// TwinCAT 3 PLC project MyLibrary_Test
// ProgramVersion: 3.1.4023.0
// libraries:
//   MyLibrary, * (FabioBolognesi)
//   TcUnit, * (www.tcunit.org)
//   Tc2_Standard, * (Beckhoff Automation GmbH)
//   Tc2_System, * (Beckhoff Automation GmbH)
//   Tc3_Module, * (Beckhoff Automation GmbH)
// project tree:
//   / PlcTask.TcTTO
//   PROGRAMs/ MAIN.TcPOU
//   TESTs/ FB_Conversion_Test.TcPOU, FB_Interpolate_Test.TcPOU, FB_Math_Test.TcPOU, FB_StringBuilder_Test.TcPOU, FB_Sweep_Test.TcPOU, FB_Timer_Test.TcPOU

CONFIGURATION MyLibrary_Test
    RESOURCE PLC ON TwinCAT3
        TASK PlcTask(INTERVAL := T#10ms, PRIORITY := 20);
        PROGRAM MAIN WITH PlcTask : MAIN;
    END_RESOURCE
END_CONFIGURATION

// ---- PROGRAMs/MAIN.TcPOU
// PROGRAMMA DEI TEST: basta dichiarare un'istanza di ogni test suite e chiamare TcUnit.RUN().
// Per aggiungere una suite: crearla in TESTs (EXTENDS TcUnit.FB_TestSuite) e dichiararla qui.
PROGRAM MAIN
VAR
	fbInterpolateTest		:	FB_Interpolate_Test;
	fbMathTest				:	FB_Math_Test;
	fbConversionTest		:	FB_Conversion_Test;
	fbTimerTest				:	FB_Timer_Test;
	fbSweepTest				:	FB_Sweep_Test;
	fbStringBuilderTest		:	FB_StringBuilder_Test;
END_VAR

TcUnit.RUN();

END_PROGRAM

// ---- TESTs/FB_Interpolate_Test.TcPOU
// TEST DI F_InterpolateReal E F_InterpolateTime
FUNCTION_BLOCK FB_Interpolate_Test EXTENDS TcUnit.FB_TestSuite
VAR
END_VAR

MidPoint();
ClampBelow();
ClampAbove();
ReversedPoints();
SamePoints();
InterpolateTime();

METHOD PRIVATE ClampAbove
TEST('ClampAbove');

AssertEquals_REAL(
	Expected	:=	100,
	Actual		:=	ML.F_InterpolateReal(rX0 := 0, rX1 := 10, rY0 := 0, rY1 := 100, rX := 20),
	Delta		:=	0.0001,
	Message		:=	'Dopo il secondo punto deve restituire rY1');

TEST_FINISHED();
END_METHOD

METHOD PRIVATE ClampBelow
TEST('ClampBelow');

AssertEquals_REAL(
	Expected	:=	0,
	Actual		:=	ML.F_InterpolateReal(rX0 := 0, rX1 := 10, rY0 := 0, rY1 := 100, rX := -5),
	Delta		:=	0.0001,
	Message		:=	'Prima del primo punto deve restituire rY0');

TEST_FINISHED();
END_METHOD

METHOD PRIVATE InterpolateTime
TEST('InterpolateTime');

AssertEquals_REAL(
	Expected	:=	2.5,
	Actual		:=	ML.F_InterpolateTime(tX0 := T#0S, tX1 := T#2S, rY0 := 0, rY1 := 10, tX := T#500MS),
	Delta		:=	0.0001,
	Message		:=	'Interpolazione con ascisse TIME');

TEST_FINISHED();
END_METHOD

METHOD PRIVATE MidPoint
TEST('MidPoint');

AssertEquals_REAL(
	Expected	:=	50,
	Actual		:=	ML.F_InterpolateReal(rX0 := 0, rX1 := 10, rY0 := 0, rY1 := 100, rX := 5),
	Delta		:=	0.0001,
	Message		:=	'Punto medio');

TEST_FINISHED();
END_METHOD

METHOD PRIVATE ReversedPoints
TEST('ReversedPoints');

AssertEquals_REAL(
	Expected	:=	25,
	Actual		:=	ML.F_InterpolateReal(rX0 := 10, rX1 := 0, rY0 := 100, rY1 := 0, rX := 2.5),
	Delta		:=	0.0001,
	Message		:=	'Punti in ordine decrescente: interpolazione');
AssertEquals_REAL(
	Expected	:=	100,
	Actual		:=	ML.F_InterpolateReal(rX0 := 10, rX1 := 0, rY0 := 100, rY1 := 0, rX := 20),
	Delta		:=	0.0001,
	Message		:=	'Punti in ordine decrescente: saturazione');

TEST_FINISHED();
END_METHOD

METHOD PRIVATE SamePoints
TEST('SamePoints');

AssertEquals_REAL(
	Expected	:=	7,
	Actual		:=	ML.F_InterpolateReal(rX0 := 3, rX1 := 3, rY0 := 7, rY1 := 9, rX := 5),
	Delta		:=	0.0001,
	Message		:=	'Con rX0 = rX1 deve restituire rY0');

TEST_FINISHED();
END_METHOD

END_FUNCTION_BLOCK

// ---- TESTs/FB_Math_Test.TcPOU
// TEST DI F_Saturation E F_Atan2
FUNCTION_BLOCK FB_Math_Test EXTENDS TcUnit.FB_TestSuite
VAR
END_VAR

Saturation();
Atan2Quadrants();

METHOD PRIVATE Atan2Quadrants
VAR
	rPi	:	REAL	:=	ML.GVL_Constants.PI;
END_VAR
TEST('Atan2Quadrants');

AssertEquals_REAL(Expected := rPi / 4,		Actual := ML.F_Atan2(rX := 1,	rY := 1),	Delta := 0.0001, Message := 'Primo quadrante');
AssertEquals_REAL(Expected := 3 * rPi / 4,	Actual := ML.F_Atan2(rX := -1,	rY := 1),	Delta := 0.0001, Message := 'Secondo quadrante');
AssertEquals_REAL(Expected := -3 * rPi / 4,	Actual := ML.F_Atan2(rX := -1,	rY := -1),	Delta := 0.0001, Message := 'Terzo quadrante');
AssertEquals_REAL(Expected := -rPi / 4,		Actual := ML.F_Atan2(rX := 1,	rY := -1),	Delta := 0.0001, Message := 'Quarto quadrante');
AssertEquals_REAL(Expected := rPi / 2,		Actual := ML.F_Atan2(rX := 0,	rY := 1),	Delta := 0.0001, Message := 'Asse Y positivo');
AssertEquals_REAL(Expected := 0,			Actual := ML.F_Atan2(rX := 0,	rY := 0),	Delta := 0.0001, Message := 'Origine');

TEST_FINISHED();
END_METHOD

METHOD PRIVATE Saturation
TEST('Saturation');

AssertEquals_REAL(Expected := 5,	Actual := ML.F_Saturation(rInput := 5,	rMinimumValue := 0, rMaximumValue := 10), Delta := 0.0001, Message := 'Valore interno');
AssertEquals_REAL(Expected := 0,	Actual := ML.F_Saturation(rInput := -3,	rMinimumValue := 0, rMaximumValue := 10), Delta := 0.0001, Message := 'Sotto il minimo');
AssertEquals_REAL(Expected := 10,	Actual := ML.F_Saturation(rInput := 12,	rMinimumValue := 0, rMaximumValue := 10), Delta := 0.0001, Message := 'Sopra il massimo');

TEST_FINISHED();
END_METHOD

END_FUNCTION_BLOCK

// ---- TESTs/FB_Conversion_Test.TcPOU
// TEST DI F_TimeToSeconds E F_SecondsToTime
FUNCTION_BLOCK FB_Conversion_Test EXTENDS TcUnit.FB_TestSuite
VAR
END_VAR

TimeToSeconds();
SecondsToTime();

METHOD PRIVATE SecondsToTime
TEST('SecondsToTime');

AssertEquals_TIME(
	Expected	:=	T#2S250MS,
	Actual		:=	ML.F_SecondsToTime(2.25),
	Message		:=	'2,25 s');

TEST_FINISHED();
END_METHOD

METHOD PRIVATE TimeToSeconds
TEST('TimeToSeconds');

AssertEquals_REAL(
	Expected	:=	1.5,
	Actual		:=	ML.F_TimeToSeconds(T#1S500MS),
	Delta		:=	0.0001,
	Message		:=	'1,5 s');

TEST_FINISHED();
END_METHOD

END_FUNCTION_BLOCK

// ---- TESTs/FB_Timer_Test.TcPOU
// TEST DI FB_Timer
FUNCTION_BLOCK FB_Timer_Test EXTENDS TcUnit.FB_TestSuite
VAR
	fbElapsed	:	ML.FB_Timer;
	fbSelf		:	ML.FB_Timer;
	fbReset		:	ML.FB_Timer;
END_VAR

VerifyElapsed();
VerifySelfElapsed();
ResetCondition();

METHOD PRIVATE ResetCondition
TEST('ResetCondition');

fbReset.ResetWithOffset(T#5S);
AssertFalse(Condition := fbReset.ResetCondition(FALSE),	Message := 'Condizione FALSE: nessun reset');
AssertTrue(Condition := fbReset.VerifyElapsed(T#4S),		Message := 'Senza reset il tempo trascorso resta 5 s');
AssertTrue(Condition := fbReset.ResetCondition(TRUE),		Message := 'Condizione TRUE: reset eseguito');
AssertFalse(Condition := fbReset.VerifyElapsed(T#1S),		Message := 'Dopo il reset il tempo riparte da 0');

TEST_FINISHED();
END_METHOD

METHOD PRIVATE VerifyElapsed
TEST('VerifyElapsed');

fbElapsed.ResetWithOffset(T#2S);
AssertTrue(Condition := fbElapsed.VerifyElapsed(T#1S),	Message := 'Sono passati 2 s: 1 s deve risultare trascorso');
AssertFalse(Condition := fbElapsed.VerifyElapsed(T#10S),	Message := 'Sono passati 2 s: 10 s non devono risultare trascorsi');

TEST_FINISHED();
END_METHOD

METHOD PRIVATE VerifySelfElapsed
TEST('VerifySelfElapsed');

fbSelf.ResetWithOffset(T#2S);
fbSelf.ChangeTimer(T#1S);
AssertTrue(Condition := fbSelf.VerifySelfElapsed(),	Message := 'Durata 1 s, trascorsi 2 s');
fbSelf.ChangeTimer(T#10S);
AssertFalse(Condition := fbSelf.VerifySelfElapsed(),	Message := 'Durata 10 s, trascorsi 2 s');

TEST_FINISHED();
END_METHOD

END_FUNCTION_BLOCK

// ---- TESTs/FB_Sweep_Test.TcPOU
// TEST DI FB_Sweep
FUNCTION_BLOCK FB_Sweep_Test EXTENDS TcUnit.FB_TestSuite
VAR
	fbInvalid	:	ML.FB_Sweep;
	fbStart		:	ML.FB_Sweep;
END_VAR

InitializeRejectsZeroDuration();
StartValues();

METHOD PRIVATE InitializeRejectsZeroDuration
TEST('InitializeRejectsZeroDuration');

AssertFalse(
	Condition	:=	fbInvalid.Initialize(rInputStartFrequency := 1, rInputEndFrequency := 10, rInputDuration := 0),
	Message		:=	'Durata nulla: Initialize deve restituire FALSE');

TEST_FINISHED();
END_METHOD

METHOD PRIVATE StartValues
TEST('StartValues');

AssertTrue(
	Condition	:=	fbStart.Initialize(rInputStartFrequency := 1, rInputEndFrequency := 10, rInputDuration := 5),
	Message		:=	'Parametri validi: Initialize deve restituire TRUE');
fbStart.Start();
// APPENA PARTITO: FREQUENZA = FREQUENZA INIZIALE E USCITA QUASI NULLA (seno di un angolo piccolo)
AssertEquals_REAL(Expected := 1,	Actual := fbStart.ComputeFrequency(),	Delta := 0.1,	Message := 'Frequenza iniziale');
AssertEquals_REAL(Expected := 0,	Actual := fbStart.Step(),				Delta := 0.1,	Message := 'Uscita iniziale');

TEST_FINISHED();
END_METHOD

END_FUNCTION_BLOCK

// ---- TESTs/FB_StringBuilder_Test.TcPOU
// TEST DI FB_StringBuilder
FUNCTION_BLOCK FB_StringBuilder_Test EXTENDS TcUnit.FB_TestSuite
VAR
	fbAddChar	:	ML.FB_StringBuilder;
	fbAddString	:	ML.FB_StringBuilder;
	fbOverflow	:	ML.FB_StringBuilder;
	fbBuild	:	ML.FB_StringBuilder;
	fbKeyValue	:	ML.FB_StringBuilder;
	fbDelete	:	ML.FB_StringBuilder;
	fbReset	:	ML.FB_StringBuilder;
	sResult	:	STRING(255);
END_VAR

AddChar();
AddString();
Overflow();
BuildString();
AddKeyValue();
DeleteChars();
ResetBuffer();

METHOD PRIVATE AddChar
TEST('AddChar');

AssertTrue(Condition := fbAddChar.AddChar(ML.E_Ascii.OpenParenthesis),	Message := 'AddChar');
AssertTrue(Condition := fbAddChar.AddByte(65),								Message := 'AddByte (A)');
AssertTrue(Condition := fbAddChar.AddChar(ML.E_Ascii.CloseParenthesis),	Message := 'AddChar');
fbAddChar.BuildString(ADR(sResult), SIZEOF(sResult));
AssertEquals_STRING(Expected := '(A)', Actual := sResult, Message := 'Contenuto');

TEST_FINISHED();
END_METHOD

METHOD PRIVATE AddKeyValue
VAR
	sKey	:	STRING	:=	'a';
	sValue	:	STRING	:=	'1';
END_VAR
TEST('AddKeyValue');

AssertTrue(Condition := fbKeyValue.AddKeyValue(ADR(sKey), ADR(sValue)),	Message := 'Chiave e valore validi');
AssertFalse(Condition := fbKeyValue.AddKeyValue(0, ADR(sValue)),			Message := 'Chiave nulla');
fbKeyValue.BuildString(ADR(sResult), SIZEOF(sResult));
AssertEquals_STRING(Expected := 'a:1,', Actual := sResult, Message := 'Contenuto');

TEST_FINISHED();
END_METHOD

METHOD PRIVATE AddString
VAR
	sText	:	STRING	:=	'ciao';
END_VAR
TEST('AddString');

AssertTrue(Condition := fbAddString.AddString(ADR(sText)),	Message := 'Stringa valida');
AssertFalse(Condition := fbAddString.AddString(0),			Message := 'Puntatore nullo');
fbAddString.BuildString(ADR(sResult), SIZEOF(sResult));
AssertEquals_STRING(Expected := 'ciao', Actual := sResult, Message := 'Contenuto');

TEST_FINISHED();
END_METHOD

METHOD PRIVATE BuildString
VAR
	sShort	:	STRING(10);
	sText	:	STRING	:=	'ciao';
	sLong	:	STRING	:=	' molto lungo';
END_VAR
TEST('BuildString');

fbBuild.AddString(ADR(sText));
AssertTrue(Condition := fbBuild.BuildString(ADR(sShort), SIZEOF(sShort)),	Message := 'Il testo entra nella destinazione');
AssertEquals_STRING(Expected := 'ciao', Actual := sShort, Message := 'Contenuto');
AssertTrue(Condition := fbBuild.BuildString(ADR(sShort), SIZEOF(sShort)),	Message := 'Seconda chiamata a BuildString');
AssertEquals_STRING(Expected := 'ciao', Actual := sShort, Message := 'Contenuto dopo la seconda chiamata');

fbBuild.AddString(ADR(sLong));
AssertFalse(Condition := fbBuild.BuildString(ADR(sShort), SIZEOF(sShort)),	Message := 'Destinazione troppo piccola');
AssertEquals_STRING(Expected := 'ciao', Actual := sShort, Message := 'La destinazione non deve essere toccata');
AssertFalse(Condition := fbBuild.BuildString(0, 100),							Message := 'Destinazione nulla');

TEST_FINISHED();
END_METHOD

METHOD PRIVATE DeleteChars
VAR
	sText	:	STRING	:=	'abc';
END_VAR
TEST('DeleteChars');

fbDelete.AddString(ADR(sText));
AssertTrue(Condition := fbDelete.DeleteChars(1),	Message := 'Cancello 1 carattere su 3');
fbDelete.BuildString(ADR(sResult), SIZEOF(sResult));
AssertEquals_STRING(Expected := 'ab', Actual := sResult, Message := 'Contenuto dopo la prima cancellazione');
AssertFalse(Condition := fbDelete.DeleteChars(5),	Message := 'Cancello 5 caratteri su 2');
fbDelete.BuildString(ADR(sResult), SIZEOF(sResult));
AssertEquals_STRING(Expected := '', Actual := sResult, Message := 'Contenuto dopo la seconda cancellazione');

TEST_FINISHED();
END_METHOD

METHOD PRIVATE Overflow
VAR
	udiCount	:	UDINT;
	bAllAdded	:	BOOL	:=	TRUE;
END_VAR
TEST('Overflow');

// IL BUFFER CONTIENE ESATTAMENTE MAX_CHARACTERS CARATTERI: IL SUCCESSIVO DEVE ESSERE RIFIUTATO
FOR udiCount := 1 TO ML.GVL_Parameters.MAX_CHARACTERS DO
	bAllAdded	:=	bAllAdded AND fbOverflow.AddChar(ML.E_Ascii.Space);
END_FOR
AssertTrue(Condition := bAllAdded,							Message := 'Buffer riempito fino al limite');
AssertFalse(Condition := fbOverflow.AddChar(ML.E_Ascii.Space),	Message := 'Buffer pieno: AddChar deve restituire FALSE');

TEST_FINISHED();
END_METHOD

METHOD PRIVATE ResetBuffer
VAR
	sText	:	STRING	:=	'abc';
END_VAR
TEST('ResetBuffer');

fbReset.AddString(ADR(sText));
fbReset.ResetBuffer();
fbReset.BuildString(ADR(sResult), SIZEOF(sResult));
AssertEquals_STRING(Expected := '', Actual := sResult, Message := 'Dopo ResetBuffer il testo deve essere vuoto');

TEST_FINISHED();
END_METHOD

END_FUNCTION_BLOCK
